              [0]
                bool bANDOR[2]
                num nSigIndex[3]
                num nSigType[3]
                num nValue[3]
            mdesc mMdesc = {leave=0}
            num nActionIndex = 60
            num nDelay = 1
            num nMoveType = 1
            num nPercentage
            num nSigValue = 1
        pointRx pPointRx[2] = {x=-431.230414, y=-162.0462365, z=907.0568155, rx=-0.848018, ry=1.454542, rz=-89.586966, shoulder=lefty, elbow=epositive, wrist=wpositive}
        string sID
      [26]
        bool bMarked
        jointRx jJointRx = {j1=-166.933303, j2=-27.00897371, j3=131.996075, j4=-179.481483, j5=106.595535, j6=257.47678}
        pointRx pInter
        paraItem pParaItem
          [0]
            bool bSafePoint
            ifItem iIfItem
              [0]
                bool bANDOR[2]
                num nSigIndex[3]
                num nSigType[3]
                num nValue[3]
            mdesc mMdesc = {leave=0}
            num nActionIndex = 60
            num nDelay = 1
            num nMoveType = 1
            num nPercentage
            num nSigValue = 1
        pointRx pPointRx[2] = {x=-478.459752, y=-121.00621071, z=907.0567925, rx=-0.848076, ry=1.454961, rz=-89.586876, shoulder=lefty, elbow=epositive, wrist=wpositive}
        string sID
      [27]
        bool bMarked
        jointRx jJointRx = {j1=-161.359654, j2=-43.128032, j3=139.566973, j4=-179.65854, j5=98.0893894, j6=251.805285}
        pointRx pInter
        paraItem pParaItem
          [0]
            bool bSafePoint
            ifItem iIfItem
              [0]
                bool bANDOR[2]
                num nSigIndex[3]
                num nSigType[3]
                num nValue[3]
            mdesc mMdesc = {leave=0}
            num nActionIndex = 60
            num nDelay = 1
            num nMoveType = 1
            num nPercentage
            num nSigValue = 1
        pointRx pPointRx[2] = {x=-370.0723683, y=-121.00622289, z=907.0568097, rx=-0.848122, ry=1.455866, rz=-89.586773, shoulder=lefty, elbow=epositive, wrist=wpositive}
        string sID
      [28]
        bool bMarked
        jointRx jJointRx = {j1=-149.438088, j2=-59.165199, j3=144.268192, j4=-180.0110509, j5=86.787986, j6=239.841608}
        pointRx pInter
        paraItem pParaItem
          [0]
            bool bSafePoint
            ifItem iIfItem
              [0]
                bool bANDOR[2]
                num nSigIndex[3]
                num nSigType[3]
                num nValue[3]
            mdesc mMdesc = {leave=0}
            num nActionIndex = 60
            num nDelay = 1
            num nMoveType = 1
            num nPercentage
            num nSigValue = 1
        pointRx pPointRx[2] = {x=-264.506872, y=-121.0396803, z=907.056801, rx=-0.847447, ry=1.456472, rz=-89.58649, shoulder=lefty, elbow=epositive, wrist=wpositive}
        string sID
      [29]
        bool bMarked
        jointRx jJointRx = {j1=-109.352401, j2=-55.463724, j3=143.190298, j4=-179.110187, j5=94.66122, j6=199.697269}
        pointRx pInter
        paraItem pParaItem
          [0]
            bool bSafePoint
            ifItem iIfItem
              [0]
                bool bANDOR[2]
                num nSigIndex[3]
                num nSigType[3]
                num nValue[3]
            mdesc mMdesc = {leave=0}
            num nActionIndex = 60
            num nDelay = 1
            num nMoveType = 1
            num nPercentage
            num nSigValue = 1
        pointRx pPointRx[2] = {x=-159.72072, y=-122.885758, z=904.993295, rx=-6.838913, ry=1.455718, rz=-89.586721, shoulder=lefty, elbow=epositive, wrist=wpositive}
        string sID
      [30]
        bool bMarked
        jointRx jJointRx = {j1=-79.892893, j2=-62.95293, j3=144.690953, j4=-181.59506, j5=82.320479, j6=170.516449}
        pointRx pInter
        paraItem pParaItem
          [0]
            bool bSafePoint
            ifItem iIfItem
              [0]
                bool bANDOR[2]
                num nSigIndex[3]
                num nSigType[3]
                num nValue[3]
            mdesc mMdesc = {leave=0}
            num nActionIndex = 60
            num nDelay = 1
            num nMoveType = 1
            num nPercentage
            num nSigValue = 1
        pointRx pPointRx[2] = {x=-69.346685, y=-130.105505, z=910.214741, rx=-0.847967, ry=1.45452, rz=-89.58688, shoulder=lefty, elbow=epositive, wrist=wpositive}
        string sID
      [31]
        bool bMarked
        jointRx jJointRx = {j1=-72.0759477, j2=-63.259281, j3=144.746667, j4=-181.66354, j5=81.850252, j6=162.71938}
        pointRx pInter
        paraItem pParaItem
          [0]
            bool bSafePoint
            ifItem iIfItem
              [0]
                bool bANDOR[2]
                num nSigIndex[3]
                num nSigType[3]
                num nValue[3]
            mdesc mMdesc = {leave=0}
            num nActionIndex = 60
            num nDelay = 1
            num nMoveType = 1
            num nPercentage
            num nSigValue = 1
        pointRx pPointRx[2] = {x=-51.755771, y=-117.0791425, z=910.214718, rx=-0.848914, ry=1.456167, rz=-89.586835, shoulder=lefty, elbow=epositive, wrist=wpositive}
        string sID
      [32]
        bool bMarked
        jointRx jJointRx = {j1=-44.811682, j2=-48.0293352, j3=140.945616, j4=-181.628999, j5=92.47994, j6=135.137458}
        pointRx pInter
        paraItem pParaItem
          [0]
            bool bSafePoint
            ifItem iIfItem
              [0]
                bool bANDOR[2]
                num nSigIndex[3]
                num nSigType[3]
                num nValue[3]
            mdesc mMdesc = {leave=0}
            num nActionIndex = 60
            num nDelay = 1
            num nMoveType = 1
            num nPercentage
            num nSigValue = 1
        pointRx pPointRx[2] = {x=51.963327, y=-117.113206, z=910.214709, rx=-0.848031, ry=1.455725, rz=-89.586763, shoulder=lefty, elbow=epositive, wrist=wpositive}
        string sID
      [33]
        bool bMarked
        jointRx jJointRx = {j1=-31.191441, j2=-31.775365, j3=134.235516, j4=-181.510713, j5=101.649355, j6=121.278415}
        pointRx pInter
        paraItem pParaItem
          [0]
            bool bSafePoint
            ifItem iIfItem
              [0]
                bool bANDOR[2]
                num nSigIndex[3]
                num nSigType[3]
                num nValue[3]
            mdesc mMdesc = {leave=0}
            num nActionIndex = 60
            num nDelay = 1
            num nMoveType = 1
            num nPercentage
            num nSigValue = 1
        pointRx pPointRx[2] = {x=158.149141, y=-117.113148, z=910.214664, rx=-0.848148, ry=1.456314, rz=-89.586714, shoulder=lefty, elbow=epositive, wrist=wpositive}
        string sID
      [34]
        bool bMarked
        jointRx jJointRx = {j1=-40.0816208, j2=-16.835573, j3=125.131891, j4=-181.666835, j5=107.718754, j6=129.975311}
        pointRx pInter
        paraItem pParaItem
          [0]
            bool bSafePoint
            ifItem iIfItem
              [0]
                bool bANDOR[2]
                num nSigIndex[3]
                num nSigType[3]
                num nValue[3]
            mdesc mMdesc = {leave=0}
            num nActionIndex = 60
            num nDelay = 1
            num nMoveType = 1
            num nPercentage
            num nSigValue = 1
        pointRx pPointRx[2] = {x=214.525801, y=-229.162911, z=909.73734, rx=-0.84777, ry=1.458696, rz=-89.580189, shoulder=lefty, elbow=epositive, wrist=wpositive}
        string sID
      [35]
        bool bMarked
        jointRx jJointRx = {j1=-38.0065024, j2=-21.286047, j3=118.71891, j4=-181.579059, j5=96.805117, j6=128.219507}
        pointRx pInter
        paraItem pParaItem
          [0]
            bool bSafePoint
            ifItem iIfItem
              [0]
                bool bANDOR[2]
                num nSigIndex[3]
                num nSigType[3]
                num nValue[3]
            mdesc mMdesc = {leave=0}
            num nActionIndex = 60
            num nDelay = 1
            num nMoveType = 1
            num nPercentage
            num nSigValue = 1
        pointRx pPointRx[2] = {x=212.211278, y=-207.646289, z=998.566722, rx=-0.850784, ry=1.457906, rz=-89.580462, shoulder=lefty, elbow=epositive, wrist=wpositive}
        string sID
      [36]
        bool bMarked
        jointRx jJointRx = {j1=-52.752521, j2=-35.622941, j3=126.84106, j4=-181.674406, j5=91.0121163, j6=143.128467}
        pointRx pInter
        paraItem pParaItem
          [0]
            bool bSafePoint
            ifItem iIfItem
              [0]
                bool bANDOR[2]
                num nSigIndex[3]
                num nSigType[3]
                num nValue[3]
            mdesc mMdesc = {leave=0}
            num nActionIndex = 60
            num nDelay = 1
            num nMoveType = 1
            num nPercentage
            num nSigValue = 1
        pointRx pPointRx[2] = {x=81.927573, y=-207.64624, z=998.566713, rx=-0.849883, ry=1.457004, rz=-89.580659, shoulder=lefty, elbow=epositive, wrist=wpositive}
        string sID
      [37]
        bool bMarked
        jointRx jJointRx = {j1=-77.0870811, j2=-46.879063, j3=131.352455, j4=-181.617077, j5=84.978132, j6=167.644391}
        pointRx pInter
        paraItem pParaItem
          [0]
            bool bSafePoint
            ifItem iIfItem
              [0]
                bool bANDOR[2]
                num nSigIndex[3]
                num nSigType[3]
                num nValue[3]
            mdesc mMdesc = {leave=0}
            num nActionIndex = 60
            num nDelay = 1
            num nMoveType = 1
            num nPercentage
            num nSigValue = 1
        pointRx pPointRx[2] = {x=-43.990353, y=-207.646288, z=998.566728, rx=-0.850075, ry=1.457778, rz=-89.580533, shoulder=lefty, elbow=epositive, wrist=wpositive}
        string sID
      [38]
        bool bMarked
        jointRx jJointRx = {j1=-111.116903, j2=-50.0659704, j3=132.355862, j4=-181.0596149, j5=83.609194, j6=201.655459}
        pointRx pInter
        paraItem pParaItem
          [0]
            bool bSafePoint
            ifItem iIfItem
              [0]
                bool bANDOR[2]
                num nSigIndex[3]
                num nSigType[3]
                num nValue[3]
            mdesc mMdesc = {leave=0}
            num nActionIndex = 60
            num nDelay = 1
            num nMoveType = 1
            num nPercentage
            num nSigValue = 1
        pointRx pPointRx[2] = {x=-174.289788, y=-207.64635, z=998.566731, rx=-0.850332, ry=1.457213, rz=-89.580703, shoulder=lefty, elbow=epositive, wrist=wpositive}
        string sID
      [39]
        bool bMarked
        jointRx jJointRx = {j1=-137.0855759, j2=-42.345518, j3=129.720085, j4=-180.369378, j5=89.0207368, j6=227.505532}
        pointRx pInter
        paraItem pParaItem
          [0]
            bool bSafePoint
            ifItem iIfItem
              [0]
                bool bANDOR[2]
                num nSigIndex[3]
                num nSigType[3]
                num nValue[3]
            mdesc mMdesc = {leave=0}
            num nActionIndex = 60
            num nDelay = 1
            num nMoveType = 1
            num nPercentage
            num nSigValue = 1
        pointRx pPointRx[2] = {x=-302.979782, y=-207.646334, z=998.566722, rx=-0.85052, ry=1.457032, rz=-89.580847, shoulder=lefty, elbow=epositive, wrist=wpositive}
        string sID
      [40]
        bool bMarked
        jointRx jJointRx = {j1=-151.0508911, j2=-29.171185, j3=123.534262, j4=-179.961205, j5=96.0495583, j6=241.462817}
        pointRx pInter
        paraItem pParaItem
          [0]
            bool bSafePoint
            ifItem iIfItem
              [0]
                bool bANDOR[2]
                num nSigIndex[3]
                num nSigType[3]
                num nValue[3]
            mdesc mMdesc = {leave=0}
            num nActionIndex = 60
            num nDelay = 1
            num nMoveType = 1
            num nPercentage
            num nSigValue = 1
        pointRx pPointRx[2] = {x=-430.862611, y=-207.646306, z=998.566713, rx=-0.850258, ry=1.457026, rz=-89.580783, shoulder=lefty, elbow=epositive, wrist=wpositive}
        string sID
      [41]
        bool bMarked
        jointRx jJointRx = {j1=-158.836736, j2=-14.491785, j3=113.841224, j4=-179.728571, j5=101.0150294, j6=249.293251}
        pointRx pInter
        paraItem pParaItem
          [0]
            bool bSafePoint
            ifItem iIfItem
              [0]
                bool bANDOR[2]
                num nSigIndex[3]
                num nSigType[3]
                num nValue[3]
            mdesc mMdesc = {leave=0}
            num nActionIndex = 60
            num nDelay = 1
            num nMoveType = 1
            num nPercentage
            num nSigValue = 1
        pointRx pPointRx[2] = {x=-562.67346, y=-207.646298, z=998.566704, rx=-0.85004, ry=1.457102, rz=-89.580664, shoulder=lefty, elbow=epositive, wrist=wpositive}
        string sID
      [42]
        bool bMarked
        jointRx jJointRx = {j1=-155.845923, j2=-13.0548146, j3=111.92039, j4=-188.865529, j5=96.422595, j6=245.198525}
        pointRx pInter
        paraItem pParaItem
          [0]
            bool bSafePoint
            ifItem iIfItem
              [0]
                bool bANDOR[2]
                num nSigIndex[3]
                num nSigType[3]
                num nValue[3]
            mdesc mMdesc = {leave=0}
            num nActionIndex = 60
            num nDelay = 1
            num nMoveType = 1
            num nPercentage
            num nSigValue = 1
        pointRx pPointRx[2] = {x=-562.638161, y=-337.888562, z=998.56672, rx=9.00287984, ry=1.457962, rz=-89.580315, shoulder=lefty, elbow=epositive, wrist=wpositive}
        string sID
      [43]
        bool bMarked
        jointRx jJointRx = {j1=-147.535096, j2=-26.82312, j3=121.400491, j4=-188.375674, j5=90.94631, j6=237.665248}
        pointRx pInter
        paraItem pParaItem
          [0]
            bool bSafePoint
            ifItem iIfItem
              [0]
                bool bANDOR[2]
                num nSigIndex[3]
                num nSigType[3]
                num nValue[3]
            mdesc mMdesc = {leave=0}
            num nActionIndex = 60
            num nDelay = 1
            num nMoveType = 1
            num nPercentage
            num nSigValue = 1
        pointRx pPointRx[2] = {x=-432.220001, y=-337.853364, z=998.566714, rx=9.00213484, ry=1.459063, rz=-89.580213, shoulder=lefty, elbow=epositive, wrist=wpositive}
        string sID
      [44]
        bool bMarked
        jointRx jJointRx = {j1=-132.698615, j2=-39.252375, j3=127.676364, j4=-187.225333, j5=82.829942, j6=223.785577}
        pointRx pInter
        paraItem pParaItem
          [0]
            bool bSafePoint
            ifItem iIfItem
              [0]
                bool bANDOR[2]
                num nSigIndex[3]
                num nSigType[3]
                num nValue[3]
            mdesc mMdesc = {leave=0}
            num nActionIndex = 60
            num nDelay = 1
            num nMoveType = 1
            num nPercentage
            num nSigValue = 1
        pointRx pPointRx[2] = {x=-300.123089, y=-337.853319, z=998.566719, rx=9.00234408, ry=1.458849, rz=-89.580203, shoulder=lefty, elbow=epositive, wrist=wpositive}
        string sID
      [45]
        bool bMarked
        jointRx jJointRx = {j1=-108.42449, j2=-45.841755, j3=130.208449, j4=-184.343765, j5=76.313958, j6=199.690032}
        pointRx pInter
        paraItem pParaItem
          [0]
            bool bSafePoint
            ifItem iIfItem
              [0]
                bool bANDOR[2]
                num nSigIndex[3]
                num nSigType[3]
                num nValue[3]
            mdesc mMdesc = {leave=0}
            num nActionIndex = 60
            num nDelay = 1
            num nMoveType = 1
            num nPercentage
            num nSigValue = 1
        pointRx pPointRx[2] = {x=-172.654258, y=-337.853312, z=998.566728, rx=9.00223206, ry=1.458726, rz=-89.580305, shoulder=lefty, elbow=epositive, wrist=wpositive}
        string sID
      [46]
        bool bMarked
        jointRx jJointRx = {j1=-78.736317, j2=-43.126447, j3=129.228824, j4=-179.671742, j5=76.98965, j6=169.222407}
        pointRx pInter
        paraItem pParaItem
          [0]
            bool bSafePoint
            ifItem iIfItem
              [0]
                bool bANDOR[2]
                num nSigIndex[3]
                num nSigType[3]
                num nValue[3]
            mdesc mMdesc = {leave=0}
            num nActionIndex = 60
            num nDelay = 1
            num nMoveType = 1
            num nPercentage
            num nSigValue = 1
        pointRx pPointRx[2] = {x=-45.447251, y=-337.853389, z=998.566726, rx=9.00199945, ry=1.458945, rz=-89.580351, shoulder=lefty, elbow=epositive, wrist=wpositive}
        string sID
      [47]
        bool bMarked
        jointRx jJointRx = {j1=-55.269987, j2=-32.727334, j3=124.635868, j4=-176.0660377, j5=83.679452, j6=145.65255}
        pointRx pInter
        paraItem pParaItem
          [0]
            bool bSafePoint
            ifItem iIfItem
              [0]
                bool bANDOR[2]
                num nSigIndex[3]
                num nSigType[3]
                num nValue[3]
            mdesc mMdesc = {leave=0}
            num nActionIndex = 60
            num nDelay = 1
            num nMoveType = 1
            num nPercentage
            num nSigValue = 1
        pointRx pPointRx[2] = {x=84.070677, y=-337.853402, z=998.566717, rx=9.00187497, ry=1.458768, rz=-89.580396, shoulder=lefty, elbow=epositive, wrist=wpositive}
        string sID
      [48]
        bool bMarked
        jointRx jJointRx = {j1=-40.841132, j2=-19.568561, j3=116.755728, j4=-174.163665, j5=90.168201, j6=131.750923}
        pointRx pInter
        paraItem pParaItem
          [0]
            bool bSafePoint
            ifItem iIfItem
              [0]
                bool bANDOR[2]
                num nSigIndex[3]
                num nSigType[3]
                num nValue[3]
            mdesc mMdesc = {leave=0}
            num nActionIndex = 60
            num nDelay = 1
            num nMoveType = 1
            num nPercentage
            num nSigValue = 1
        pointRx pPointRx[2] = {x=211.980606, y=-337.853391, z=998.566708, rx=9.00196014, ry=1.458665, rz=-89.58043, shoulder=lefty, elbow=epositive, wrist=wpositive}
        string sID
      [49]
        bool bMarked
        jointRx jJointRx = {j1=-42.435689, j2=-17.531711, j3=114.153967, j4=-181.618637, j5=96.115044, j6=132.665436}
        pointRx pInter
        paraItem pParaItem
          [0]
            bool bSafePoint
            ifItem iIfItem
              [0]
                bool bANDOR[2]
                num nSigIndex[3]
                num nSigType[3]
                num nValue[3]
            mdesc mMdesc = {leave=0}
            num nActionIndex = 60
            num nDelay = 1
            num nMoveType = 1
            num nPercentage
            num nSigValue = 1
        pointRx pPointRx[2] = {x=218.0171948, y=-256.0900536, z=1017.17652, rx=-0.847487, ry=1.458394, rz=-89.579905, shoulder=lefty, elbow=epositive, wrist=wpositive}
        string sID
      [50]
        bool bMarked
        jointRx jJointRx = {j1=-55.762863, j2=-3.783808, j3=100.0532234, j4=-191.228362, j5=109.160387, j6=143.472454}
        pointRx pInter
        paraItem pParaItem
          [0]
            bool bSafePoint
            ifItem iIfItem
              [0]
                bool bANDOR[2]
                num nSigIndex[3]
                num nSigType[3]
                num nValue[3]
            mdesc mMdesc = {leave=0}
            num nActionIndex = 60
            num nDelay = 1
            num nMoveType = 1
            num nPercentage
            num nSigValue = 1
        pointRx pPointRx[2] = {x=213.807346, y=-264.112451, z=1017.176406, rx=-16.836873, ry=1.457256, rz=-89.580052, shoulder=lefty, elbow=epositive, wrist=wpositive}
        string sID
      [51]
        bool bMarked
        jointRx jJointRx = {j1=-68.596641, j2=-12.456355, j3=107.607632, j4=-187.920513, j5=110.191419, j6=157.0455023}
        pointRx pInter
        paraItem pParaItem
          [0]
            bool bSafePoint
            ifItem iIfItem
              [0]
                bool bANDOR[2]
                num nSigIndex[3]
                num nSigType[3]
                num nValue[3]
            mdesc mMdesc = {leave=0}
            num nActionIndex = 60
            num nDelay = 1
            num nMoveType = 1
            num nPercentage
            num nSigValue = 1
        pointRx pPointRx[2] = {x=80.650673, y=-264.11245, z=1017.176424, rx=-16.836304, ry=1.456605, rz=-89.5804, shoulder=lefty, elbow=epositive, wrist=wpositive}
        string sID
      [52]
        bool bMarked
        jointRx jJointRx = {j1=-83.808916, j2=-17.800495, j3=111.680418, j4=-183.456899, j5=110.438622, j6=173.276997}
        pointRx pInter
        paraItem pParaItem
          [0]
            bool bSafePoint
            ifItem iIfItem
              [0]
                bool bANDOR[2]
                num nSigIndex[3]
                num nSigType[3]
                num nValue[3]
            mdesc mMdesc = {leave=0}
            num nActionIndex = 60
            num nDelay = 1
            num nMoveType = 1
            num nPercentage
            num nSigValue = 1
        pointRx pPointRx[2] = {x=-46.894414, y=-264.112449, z=1017.176424, rx=-16.836228, ry=1.456863, rz=-89.580298, shoulder=lefty, elbow=epositive, wrist=wpositive}
        string sID
      [53]
        bool bMarked
        jointRx jJointRx = {j1=-100.312543, j2=-19.0224916, j3=112.550808, j4=-178.360867, j5=110.350071, j6=190.859412}
        pointRx pInter
        paraItem pParaItem
          [0]
            bool bSafePoint
            ifItem iIfItem
              [0]
                bool bANDOR[2]
                num nSigIndex[3]
                num nSigType[3]
                num nValue[3]
            mdesc mMdesc = {leave=0}
            num nActionIndex = 60
            num nDelay = 1
            num nMoveType = 1
            num nPercentage
            num nSigValue = 1
        pointRx pPointRx[2] = {x=-173.546019, y=-264.112435, z=1017.176424, rx=-16.836301, ry=1.456918, rz=-89.580312, shoulder=lefty, elbow=epositive, wrist=wpositive}
        string sID
      [54]
        bool bMarked
        jointRx jJointRx = {j1=-115.98199, j2=-15.735762, j3=110.158596, j4=-173.640472, j5=110.14502, j6=207.553211}
        pointRx pInter
        paraItem pParaItem
          [0]
            bool bSafePoint
            ifItem iIfItem
              [0]
                bool bANDOR[2]
                num nSigIndex[3]
                num nSigType[3]
                num nValue[3]
            mdesc mMdesc = {leave=0}
            num nActionIndex = 60
            num nDelay = 1
            num nMoveType = 1
            num nPercentage
            num nSigValue = 1
        pointRx pPointRx[2] = {x=-302.472979, y=-264.112438, z=1017.176424, rx=-16.836265, ry=1.456899, rz=-89.580364, shoulder=lefty, elbow=epositive, wrist=wpositive}
        string sID
      [55]
        bool bMarked
        jointRx jJointRx = {j1=-128.792616, j2=-8.69318, j3=104.475144, j4=-170.118674, j5=109.679904, j6=221.195478}
        pointRx pInter
        paraItem pParaItem
          [0]
            bool bSafePoint
            ifItem iIfItem
              [0]
                bool bANDOR[2]
                num nSigIndex[3]
                num nSigType[3]
                num nValue[3]
            mdesc mMdesc = {leave=0}
            num nActionIndex = 60
            num nDelay = 1
            num nMoveType = 1
            num nPercentage
            num nSigValue = 1
        pointRx pPointRx[2] = {x=-432.523171, y=-264.112458, z=1017.176411, rx=-16.836073, ry=1.456713, rz=-89.580423, shoulder=lefty, elbow=epositive, wrist=wpositive}
        string sID
      [56]
        bool bMarked
        jointRx jJointRx = {j1=-138.261544, j2=0.587068, j3=95.793725, j4=-167.880774, j5=108.465635, j6=231.0964901}
        pointRx pInter
        paraItem pParaItem
          [0]
            bool bSafePoint
            ifItem iIfItem
              [0]
                bool bANDOR[2]
                num nSigIndex[3]
                num nSigType[3]
                num nValue[3]
            mdesc mMdesc = {leave=0}
            num nActionIndex = 60
            num nDelay = 1
            num nMoveType = 1
            num nPercentage
            num nSigValue = 1
        pointRx pPointRx[2] = {x=-560.410604, y=-264.112428, z=1017.176386, rx=-16.835778, ry=1.455682, rz=-89.580765, shoulder=lefty, elbow=epositive, wrist=wpositive}
        string sID
      [57]
        bool bMarked
        jointRx jJointRx = {j1=-137.570299, j2=7.199857, j3=101.459775, j4=-171.647292, j5=117.25334, j6=231.115547}
        pointRx pInter
        paraItem pParaItem
          [0]
            bool bSafePoint
            ifItem iIfItem
              [0]
                bool bANDOR[2]
                num nSigIndex[3]
                num nSigType[3]
                num nValue[3]
            mdesc mMdesc = {leave=0}
            num nActionIndex = 60
            num nDelay = 1
            num nMoveType = 1
            num nPercentage
            num nSigValue = 1
        pointRx pPointRx[2] = {x=-578.753869, y=-345.929429, z=912.204286, rx=-11.433753, ry=1.454925, rz=-89.581005, shoulder=lefty, elbow=epositive, wrist=wpositive}
        string sID
      [58]
        bool bMarked
        jointRx jJointRx = {j1=-55.213058, j2=3.467821, j3=105.525268, j4=-188.670392, j5=117.327621, j6=142.0620183}
        pointRx pInter
        paraItem pParaItem
          [0]
            bool bSafePoint
            ifItem iIfItem
              [0]
                bool bANDOR[2]
                num nSigIndex[3]
                num nSigType[3]
                num nValue[3]
            mdesc mMdesc = {leave=0}
            num nActionIndex = 60
            num nDelay = 1
            num nMoveType = 1
            num nPercentage
            num nSigValue = 1
        pointRx pPointRx[2] = {x=238.850933, y=-345.929349, z=912.204253, rx=-11.433611, ry=1.455813, rz=-89.580616, shoulder=lefty, elbow=epositive, wrist=wpositive}
        string sID
      [59]
        bool bMarked
        jointRx jJointRx = {j1=-39.877322, j2=0.797114, j3=105.0689975, j4=-172.877124, j5=113.430642, j6=132.7102}
        pointRx pInter
        paraItem pParaItem
          [0]
            bool bSafePoint
            ifItem iIfItem
              [0]
                bool bANDOR[2]
                num nSigIndex[3]
                num nSigType[3]
                num nValue[3]
            mdesc mMdesc = {leave=0}
            num nActionIndex = 60
            num nDelay = 1
            num nMoveType = 1
            num nPercentage
            num nSigValue = 1
        pointRx pPointRx[2] = {x=218.979943, y=-339.519997, z=912.204287, rx=0.0970883, ry=-10.105192, rz=-89.561555, shoulder=lefty, elbow=epositive, wrist=wpositive}
        string sID
      [60]
        bool bMarked
        jointRx jJointRx = {j1=-139.351675, j2=-14.308765, j3=118.506559, j4=-173.468727, j5=96.392889, j6=230.952534}
        pointRx pInter
        paraItem pParaItem
          [0]
            bool bSafePoint
            ifItem iIfItem
              [0]
                bool bANDOR[2]
                num nSigIndex[3]
                num nSigType[3]
                num nValue[3]
            mdesc mMdesc = {leave=0}
            num nActionIndex = 60
            num nDelay = 1
            num nMoveType = 1
            num nPercentage
            num nSigValue = 1
        pointRx pPointRx[2] = {x=-578.952622, y=-339.519943, z=912.204249, rx=0.0970317, ry=-10.105966, rz=-89.561786, shoulder=lefty, elbow=epositive, wrist=wpositive}
        string sID
      [61]
        bool bMarked
        jointRx jJointRx = {j1=-153.527112, j2=10.829763, j3=100.476107, j4=-187.881335, j5=124.0989587, j6=240.245027}
        pointRx pInter
        paraItem pParaItem
          [0]
            bool bSafePoint
            ifItem iIfItem
              [0]
                bool bANDOR[2]
                num nSigIndex[3]
                num nSigType[3]
                num nValue[3]
            mdesc mMdesc = {leave=0}
            num nActionIndex = 60
            num nDelay = 1
            num nMoveType = 1
            num nPercentage
            num nSigValue = 1
        pointRx pPointRx[2] = {x=-569.279809, y=-339.519992, z=912.204282, rx=0.0985985, ry=14.558774, rz=-89.603311, shoulder=lefty, elbow=epositive, wrist=wpositive}
        string sID
      [62]
        bool bMarked
        jointRx jJointRx = {j1=-64.285602, j2=-20.0957166, j3=129.0123612, j4=-193.347744, j5=102.0746215, j6=151.107564}
        pointRx pInter
        paraItem pParaItem
          [0]
            bool bSafePoint
            ifItem iIfItem
              [0]
                bool bANDOR[2]
                num nSigIndex[3]
                num nSigType[3]
                num nValue[3]
            mdesc mMdesc = {leave=0}
            num nActionIndex = 60
            num nDelay = 1
            num nMoveType = 1
            num nPercentage
            num nSigValue = 1
        pointRx pPointRx[2] = {x=213.915317, y=-339.51997, z=912.204283, rx=0.0987236, ry=14.558616, rz=-89.603162, shoulder=lefty, elbow=epositive, wrist=wpositive}
        string sID
      [63]
        bool bMarked
        jointRx jJointRx = {j1=-53.566196, j2=-35.179254, j3=137.506536, j4=-191.631372, j5=93.410669, j6=142.373056}
        pointRx pInter
        paraItem pParaItem
          [0]
            bool bSafePoint
            ifItem iIfItem
              [0]
                bool bANDOR[2]
                num nSigIndex[3]
                num nSigType[3]
                num nValue[3]
            mdesc mMdesc = {leave=0}
            num nActionIndex = 60
            num nDelay = 1
            num nMoveType = 1
            num nPercentage
            num nSigValue = 1
        pointRx pPointRx[2] = {x=213.915326, y=-213.236458, z=912.204287, rx=0.0979934, ry=14.558755, rz=-89.602991, shoulder=lefty, elbow=epositive, wrist=wpositive}
        string sID
      [64]
        bool bMarked
        jointRx jJointRx = {j1=-165.0586665, j2=8.078844, j3=103.668573, j4=-184.692599, j5=125.717529, j6=253.194344}
        pointRx pInter
        paraItem pParaItem
          [0]
            bool bSafePoint
            ifItem iIfItem
              [0]
                bool bANDOR[2]
                num nSigIndex[3]
                num nSigType[3]
                num nValue[3]
            mdesc mMdesc = {leave=0}
            num nActionIndex = 60
            num nDelay = 1
            num nMoveType = 1
            num nPercentage
            num nSigValue = 1
        pointRx pPointRx[2] = {x=-600.940306, y=-213.212092, z=912.204219, rx=0.0989693, ry=14.557609, rz=-89.603294, shoulder=lefty, elbow=epositive, wrist=wpositive}
        string sID
      [65]
        bool bMarked
        jointRx jJointRx = {j1=-153.484724, j2=-25.585659, j3=126.92235, j4=-176.190756, j5=93.457282, j6=244.405675}
        pointRx pInter
        paraItem pParaItem
          [0]
            bool bSafePoint
            ifItem iIfItem
              [0]
                bool bANDOR[2]
                num nSigIndex[3]
                num nSigType[3]
                num nValue[3]
            mdesc mMdesc = {leave=0}
            num nActionIndex = 60
            num nDelay = 1
            num nMoveType = 1
            num nPercentage
            num nSigValue = 1
        pointRx pPointRx[2] = {x=-561.0183103, y=-213.592411, z=911.589458, rx=0.0967515, ry=-8.736241, rz=-89.563414, shoulder=lefty, elbow=epositive, wrist=wpositive}
        string sID
      [66]
        bool bMarked
        jointRx jJointRx = {j1=-28.548549, j2=-4.973926, j3=111.371301, j4=-175.351676, j5=113.969198, j6=120.585782}
        pointRx pInter
        paraItem pParaItem
          [0]
            bool bSafePoint
            ifItem iIfItem
              [0]
                bool bANDOR[2]
                num nSigIndex[3]
                num nSigType[3]
                num nValue[3]
            mdesc mMdesc = {leave=0}
            num nActionIndex = 60
            num nDelay = 1
            num nMoveType = 1
            num nPercentage
            num nSigValue = 1
        pointRx pPointRx[2] = {x=243.943786, y=-213.59237, z=911.589399, rx=0.096756, ry=-8.736005, rz=-89.563446, shoulder=lefty, elbow=epositive, wrist=wpositive}
        string sID
      [67]
        bool bMarked
        jointRx jJointRx = {j1=-40.582486, j2=-11.894877, j3=121.164921, j4=-183.150746, j5=109.611524, j6=129.918427}
        pointRx pInter
        paraItem pParaItem
          [0]
            bool bSafePoint
            ifItem iIfItem
              [0]
                bool bANDOR[2]
                num nSigIndex[3]
                num nSigType[3]
                num nValue[3]
            mdesc mMdesc = {leave=0}
            num nActionIndex = 60
            num nDelay = 1
            num nMoveType = 1
            num nPercentage
            num nSigValue = 1
        pointRx pPointRx[2] = {x=243.886499, y=-240.132648, z=911.589459, rx=-2.494433, ry=1.650255, rz=-89.579218, shoulder=lefty, elbow=epositive, wrist=wpositive}
        string sID
      [68]
        bool bMarked
        jointRx jJointRx = {j1=-154.853411, j2=-5.565711, j3=115.762818, j4=-178.312294, j5=112.742312, j6=245.856073}
        pointRx pInter
        paraItem pParaItem
          [0]
            bool bSafePoint
            ifItem iIfItem
              [0]
                bool bANDOR[2]
                num nSigIndex[3]
                num nSigType[3]
                num nValue[3]
            mdesc mMdesc = {leave=0}
            num nActionIndex = 60
            num nDelay = 1
            num nMoveType = 1
            num nPercentage
            num nSigValue = 1
        pointRx pPointRx[2] = {x=-590.0361404, y=-240.107985, z=911.58941, rx=-2.495147, ry=1.649301, rz=-89.579324, shoulder=lefty, elbow=epositive, wrist=wpositive}
        string sID
      [69]
        bool bMarked
        jointRx jJointRx = {j1=-169.544974, j2=-34.564516, j3=135.652231, j4=-196.70666, j5=98.242514, j6=256.952537}
        pointRx pInter
        paraItem pParaItem
          [0]
            bool bSafePoint
            ifItem iIfItem
              [0]
                bool bANDOR[2]
                num nSigIndex[3]
                num nSigType[3]
                num nValue[3]
            mdesc mMdesc = {leave=0}
            num nActionIndex = 60
            num nDelay = 1
            num nMoveType = 1
            num nPercentage
            num nSigValue = 1
        pointRx pPointRx[2] = {x=-445.474256, y=-277.981159, z=882.163294, rx=16.699071, ry=0.613858, rz=-89.857323, shoulder=lefty, elbow=epositive, wrist=wpositive}
        string sID
      [70]
        bool bMarked
        jointRx jJointRx = {j1=-177.391687, j2=-26.280383, j3=131.71858, j4=-178.98543, j5=106.238273, j6=267.807144}
        pointRx pInter
        paraItem pParaItem
          [0]
            bool bSafePoint
            ifItem iIfItem
              [0]
                bool bANDOR[2]
                num nSigIndex[3]
                num nSigType[3]
                num nValue[3]
            mdesc mMdesc = {leave=0}
            num nActionIndex = 60
            num nDelay = 1
            num nMoveType = 1
            num nPercentage
            num nSigValue = 1
        pointRx pPointRx[2] = {x=-508.182047, y=-56.0714362, z=903.88543, rx=-1.00968978, ry=0.757209, rz=-89.854782, shoulder=lefty, elbow=epositive, wrist=wpositive}
        string sID
      [71]
        bool bMarked
        jointRx jJointRx = {j1=-178.386803, j2=-23.774985, j3=123.0997568, j4=-178.221653, j5=99.246712, j6=269.348916}
        pointRx pInter
        paraItem pParaItem
          [0]
            bool bSafePoint
            ifItem iIfItem
              [0]
                bool bANDOR[2]
                num nSigIndex[3]
                num nSigType[3]
                num nValue[3]
            mdesc mMdesc = {leave=0}
            num nActionIndex = 60
            num nDelay = 1
            num nMoveType = 1
            num nPercentage
            num nSigValue = 1
        pointRx pPointRx[2] = {x=-550.87351, y=-44.532859, z=967.883245, rx=-1.752465, ry=-0.123022, rz=-89.326741, shoulder=lefty, elbow=epositive, wrist=wpositive}
        string sID
      [72]
        bool bMarked
        jointRx jJointRx = {j1=-177.679059, j2=-40.775255, j3=131.836988, j4=-178.243692, j5=91.0106442, j6=268.385946}
        pointRx pInter
        paraItem pParaItem
          [0]
            bool bSafePoint
            ifItem iIfItem
              [0]
                bool bANDOR[2]
                num nSigIndex[3]
                num nSigType[3]
                num nValue[3]
            mdesc mMdesc = {leave=0}
            num nActionIndex = 60
            num nDelay = 1
            num nMoveType = 1
            num nPercentage
            num nSigValue = 1
        pointRx pPointRx[2] = {x=-432.372199, y=-44.56903, z=967.883219, rx=-1.752547, ry=-0.121652, rz=-89.326737, shoulder=lefty, elbow=epositive, wrist=wpositive}
        string sID
      [73]
        bool bMarked
        jointRx jJointRx = {j1=-175.615752, j2=-61.311831, j3=137.808504, j4=-178.193576, j5=76.515805, j6=265.869398}
        pointRx pInter
        paraItem pParaItem
          [0]
            bool bSafePoint
            ifItem iIfItem
              [0]
                bool bANDOR[2]
                num nSigIndex[3]
                num nSigType[3]
                num nValue[3]
            mdesc mMdesc = {leave=0}
            num nActionIndex = 60
            num nDelay = 1
            num nMoveType = 1
            num nPercentage
            num nSigValue = 1
        pointRx pPointRx[2] = {x=-303.185709, y=-44.569005, z=967.883227, rx=-1.752444, ry=-0.121634, rz=-89.326671, shoulder=lefty, elbow=epositive, wrist=wpositive}
        string sID
      [74]
        bool bMarked
        jointRx jJointRx = {j1=-120.101249, j2=-78.704971, j3=139.88333, j4=-178.891628, j5=62.637529, j6=210.254495}
        pointRx pInter
        paraItem pParaItem
          [0]
            bool bSafePoint
            ifItem iIfItem
